// RUN: sclang-gen --emit=mlir-std %s | FileCheck %s

// CHECK-LABEL: func.func @f
// CHECK:         memref.alloca() : memref<6xi8>
// CHECK:         memref.copy
// CHECK:         memref.reinterpret_cast {{%[a-z_0-9]+}} to offset: [0], sizes: [2]
function f : int
var_input
  a : struct
    a1 : int;
    a2 : real;
  end_struct;
end_var
begin
  f := a.a1;
end_function
